FUNCTION_BLOCK FB_MotorReset
VAR_INPUT
	bResetX	:	BOOL;
	bResetY	:	BOOL;
	bResetZ	:	BOOL;
END_VAR
VAR_OUTPUT
	bReset	: BOOL := FALSE;
END_VAR
VAR_IN_OUT
	motX:	AXIS_REF;
	motY:	AXIS_REF;
	motZ:	AXIS_REF;
END_VAR
VAR
	MC_RESET_X	:	MC_RESET;
	MC_RESET_Y	:	MC_RESET;
	MC_RESET_Z	:	MC_RESET;
	
	Done_X	:	BOOL;
	Done_Y	:	BOOL;
	Done_Z	:	BOOL;
END_VAR

MC_RESET_X(
	Axis	:=	motX,
	Execute	:=	bResetX,
	Done	=>	Done_X);
	
MC_RESET_Y(
	Axis	:=	motY,
	Execute	:=	bResetY,
	Done	=>	Done_Y);
	
MC_RESET_Z(
	Axis	:=	motZ,
	Execute	:=	bResetZ,
	Done	=>	Done_Z);
	
	
IF bResetX OR bResetY OR bResetZ THEN
	bReset	:=	
		((NOT bResetX) OR Done_X) AND
		((NOT bResetY) OR Done_Y) AND
		((NOT bResetZ) OR Done_Z);
ELSE
	bReset	:=	TRUE; ///
END_IF

END_FUNCTION_BLOCK

(* stored: Version 1.1.0.1, ProductVersion 3.1.4024.15
   POU FB_MotorReset: Id {da498e27-6e66-48cb-a43c-531711c64104}, SpecialFunc None *)
